(* IEC 61131-3 sources: teller/JD_Teller_LC2_V11/Class/SafetyManager (part 3) *)

            exit;
          end_if;

          pHelpManaging := pHelpManaging^.pNext;
        end_while;
      end_if;

      pHelpPdo := pHelpPdo^.pNext;
    end_while;

    pHelpConfig := pHelpConfig^.pNext;
  end_while;

END_FUNCTION

FUNCTION VIRTUAL SafetyManager::GetThisViaServerName
	VAR_INPUT
		pObjectDotServer 	: ^CHAR;
	END_VAR
	VAR_OUTPUT
		ThisPtr 	: pVoid;
	END_VAR
  VAR
    ChannelMode : CHMODE;
  END_VAR

  ThisPtr := NIL;

  if pObjectDotServer = NIL then
    return;
  end_if;

  // get thispointer to server via name
  ChannelMode := _LookUpEmbed_C(pObjectDotServer, #ThisPtr, NIL);

  // check if it's a server
  case ChannelMode of
    _CH_CMD,
    _CH_SVR:

  else
    ThisPtr := NIL;
    LogError(e_msg:="(SafetyManager::GetThisViaServerName) Couldn't get thispointer of server:");
    LogError(e_msg:=pObjectDotServer);
  end_case;

END_FUNCTION

FUNCTION SafetyManager::GetNewMovDO
	VAR_OUTPUT
		Index 	: INT;
	END_VAR
//  VAR
//  	sd_retval : DINT;
//  END_VAR

  Index := -1;

  if CopyCmdsUsed < MAX_PDO_COPY_CMDS then
    // check if there is one available but not used
    if CopyCmdsUsed < CopyCmdsAvailable then
      Index := CopyCmdsUsed;
      CopyCmdsUsed += 1;
    else
      // we have to create a new one

(*
// connection to varan manager required
      // add data object to copy our data
      sd_retval := pVaranManager^.AddMovDO(ud_dol_type:=VARAN_DOL_ISO
                                         , p_ud_handle:=(#aCopyCmds[CopyCmdsAvailable].pHandle)$^UDINT
                                         , p_ud_MovSettings:=( #aCopyCmds[CopyCmdsAvailable].pSettings)$^UDINT
                                         , ud_type := VM_PRIORITY_2
                                         );

      //look for an error
      if ( sd_retval <> 0 ) then
        ClassState := -9;
        LogError("(SafetyManager::GetNewMovDO) Failed to add a new copy command to the VaranManager!");
        return;
      end_if;
*)
      aCopyCmds[CopyCmdsAvailable].b_Ready4Action := FALSE;

      Index := CopyCmdsAvailable;

      CopyCmdsAvailable += 1;
      CopyCmdsUsed += 1;
    end_if;
  else
    LogError("Maximum of possible PDO copy commands reached!");
  end_if;

END_FUNCTION

FUNCTION SafetyManager::CheckCPUConfigs
	VAR_OUTPUT
		ConfigsOK 	: BOOL;
	END_VAR
  VAR
  	pHelpManaging   : ^t_ManagingComponent;
    pSourceManaging : ^t_ManagingComponent;
    pHelpConfig     : ^t_CfgListElem;
    pHelpPdo        : ^t_PdoListElem;
    pLastPdo        : ^t_PdoListElem;
    IsSource        : DINT;
    PDOCount : UDINT;
  END_VAR

  // before we go into the usual check routine, we have to ensure that we have enough virtual PDOs for writing interface frames (config holds a broadcast and we have to look for possible target modules)
  CreateVirtualPDOs();

  // initialize with true (normal case is that everything is ok => now we check for errors)
  ConfigsOK := TRUE;

  PDOCount := 0;

  // check if all non-optional modules are available and all corresponding domain managing module are synchron (if necessary)
  pHelpConfig := pConfigs;
  while pHelpConfig do
    pLastPdo := NIL;
    pHelpPdo := pHelpConfig^.pFirstPdoCfg;
    while pHelpPdo do
      // if it's an interface frame and no broadcast frame
      if pHelpPdo^.PdoInfo.Info.IsInterfacePDO then
        if (pHelpPdo^.PdoInfo.Info.IFBroadCast = FALSE) then

          // check if we have already added the domain interface to the IF List
          IsSource := -1; // -1 = not found, 0 = destination, 1 = source
          pSourceManaging := NIL;
          pHelpManaging := pFirstManagingInterfaceComponent;
          while pHelpManaging do
            // if source or destination of the PDO matches our managing module path => it's an interface frame to/from this domain
            if (To_StdLib.MemCmp(pHelpManaging^.pModulePath, pHelpPdo^.PdoInfo.pSourcePath, pHelpPdo^.PdoInfo.SourcePathLen) = 0) then
              pSourceManaging := pHelpManaging;
              IsSource := 1;
              exit;
            elsif (To_StdLib.MemCmp(pHelpManaging^.pModulePath, pHelpPdo^.PdoInfo.pDestPath, pHelpPdo^.PdoInfo.DestPathLen) = 0) then
              IsSource := 0;
              exit;
            end_if;

            pHelpManaging := pHelpManaging^.pNext;
          end_while;

          // if we got a source managing module and it isn't synchron
          if pSourceManaging then
            // if this pdo is not optional => the source module also isn't
            if pHelpPdo^.PdoInfo.Info.IsOptional = FALSE then
              pSourceManaging^.InfoBits.IsOptional := FALSE;
            end_if;

            if (pSourceManaging^.InfoBits.IsSynchron = FALSE) then
              if pHelpPdo^.PdoInfo.Info.IsOptional then
                // ignore it
  //              LogError("Info: Optional interface frame can't be received, because source domain is not connected or not synchron");

                // remove the PDO from the list (if not the receiver module would wait endless for the PDO and we can't send the set bus ready to quit errors of local PDOs)
                if pLastPdo then
                  // if we had already a PDO before in this configuration we have to skip the removed PDO with the next pointer
                  pLastPdo^.pNext := pHelpPdo^.pNext;

                  To_StdLib.Free(pHelpPdo^.PdoInfo.pSourcePath);
                  To_StdLib.Free(pHelpPdo^.PdoInfo.pDestPath);
                  To_StdLib.Free(pHelpPdo);

                  pHelpPdo := pLastPdo;
                else
                  // if it was the first PDO, we have to correct the first pointer
                  pHelpConfig^.pFirstPdoCfg := pHelpPdo^.pNext;

                  To_StdLib.Free(pHelpPdo^.PdoInfo.pSourcePath);
                  To_StdLib.Free(pHelpPdo^.PdoInfo.pDestPath);
                  To_StdLib.Free(pHelpPdo);

                  pHelpPdo := pHelpConfig^.pFirstPdoCfg;
                end_if;

                if pHelpPdo = NIL then
                  exit;
                end_if;
              else
                // non-optional interface frame domain missing => error
                LogError("ERROR! Non-Optional interface frame can't be received, because domain is not connected");
                ConfigsOK := FALSE;
                ClassState := -10;
              end_if;
            end_if;
          end_if;
        end_if;
      end_if;

      PDOCount += 1;

      pLastPdo := pHelpPdo;
      pHelpPdo := pHelpPdo^.pNext;
    end_while;

    pHelpConfig := pHelpConfig^.pNext;
  end_while;

  // if now PDOs found => reset the act ID to show that there are none
  if PDOCount = 0 then
    ActPDO_ID := 0;
  end_if;

END_FUNCTION

FUNCTION SafetyManager::RemoveLocalCPUCfg
	VAR_INPUT
		SafetyNumber 	: HDINT;
	END_VAR
  VAR
  	pHelpCfg    : ^t_LocalCfgListElem;
    i : UDINT;
  END_VAR

  if LocalCPUCfgNo then
    pHelpCfg := pFirstLocalCPUCfg;
    for i := 0 to (LocalCPUCfgNo-1) do
      if pHelpCfg^.SafetyNbr = SafetyNumber then
        // found it => deactivate it
        pHelpCfg^.ConfigSize := 0;
        pHelpCfg^.ConfigSent2Master := FALSE;
        exit;
      end_if;

      pHelpCfg := pHelpCfg^.pNext;
    end_for;
  end_if;

END_FUNCTION

FUNCTION SafetyManager::ClearRoutingInformations
  VAR
  	MyPara : CmdStruct;
    MyResult : results;
    pHelpManaging : ^t_ManagingComponent;
    i : UDINT;
    pHelpCfg      : ^t_LocalCfgListElem;
  END_VAR

  // we're flushin our stuff here

  // reset number of memorized safe cpu numbers
  SafeCPU_Nbr_No := 0;

  // set ID to zero for the next mapping assignment
  ActPDO_ID := 0;

  // reset interface frameno
  InterfaceFrameNo := 0;

  // reset local interface frameno
  LocalIFNo := 0;

  // clear configurations of safety-cpus
  FreeCfgLists();

  // clear number of copy DOs used
  CopyCmdsUsed := 0;

  // reset memory usage for isochronous transfer (the values are set when distributing the PDOs)
  MyPara.aPara[0] := 0;
  pHelpManaging := pFirstManagingInterfaceComponent;
  while pHelpManaging do
    pHelpManaging^.PDOReadMemUsed := 0;
    pHelpManaging^.PDOWriteMemUsed := 0;

    MyPara.uiCmd := CMD_SM_PDO_MEM_USAGE_WR;
    pHelpManaging^.pThis^.NewInst(#MyPara, #MyResult);

    MyPara.uiCmd := CMD_SM_PDO_MEM_USAGE_RD;
    pHelpManaging^.pThis^.NewInst(#MyPara, #MyResult);

    pHelpManaging^.InfoBits.HasBeenFlushed      := FALSE;
    pHelpManaging^.InfoBits.NewTimeSyncPossible := FALSE;
    pHelpManaging^.InfoBits.SubDomainsSynchron  := FALSE;
    pHelpManaging^.InfoBits.GotIFInfo           := FALSE;
    pHelpManaging^.InfoBits.LocalConfigReady    := FALSE;
    pHelpManaging^.InfoBits.IsOptional          := TRUE;  // initialize with true, later in the init process (CheckCPUConfigs) it's checked and corrected if necessary
    // synchron bit is already true at this time (or the timeout has expired)

    pHelpManaging^.DomainNr := 16#FF;

    pHelpManaging^.SubDomainsUsed := 0;
    _memset(dest:=#pHelpManaging^.SubDomainNr, usByte:=16#FF, cntr:=sizeof(pHelpManaging^.SubDomainNr));

    pHelpManaging^.ModuleNo := 0;
    _memset(dest:=#pHelpManaging^.ModuleInfo, usByte:=16#00, cntr:=sizeof(pHelpManaging^.ModuleInfo));

    pHelpManaging := pHelpManaging^.pNext;
  end_while;

  // all local cpu configs have to be sent again on reconnect
  if LocalCPUCfgNo then
    pHelpCfg := pFirstLocalCPUCfg;
    for i := 0 to (LocalCPUCfgNo-1) do
      pHelpCfg^.ConfigSent2Master := FALSE;

      pHelpCfg := pHelpCfg^.pNext;
    end_for;
  end_if;

END_FUNCTION

FUNCTION SafetyManager::CheckPDORecycle
	VAR_INPUT
		SourceDest 	: t_SourceDest;
		pNewPDO 	: ^t_PDOElement;
	END_VAR
	VAR_OUTPUT
		pRecyclePDO 	: ^t_PDOElement;
	END_VAR
  VAR
  	i : UDINT;
    pHelpInfo : ^t_PDOModuleInfo;
    pSearchInfo : ^t_PDOModuleInfo;
    ppHelpManaging : ^t_pManagingComponent;
    pSearchManaging : ^t_ManagingComponent;
  END_VAR

  // initialize with invalid
  pRecyclePDO := NIL;

  // if we have no pdoelements yet, quit
  if PDOElementNo = 0 then
    return;
  end_if;

  // we search for a PDO with the same source (then it contains the same data)
  pHelpInfo := #aPDOElements[0].SourceInfo;
  pSearchInfo := #pNewPDO^.SourceInfo;

  case SourceDest of
    SourceDest_IsSource:
      ppHelpManaging := #aPDOElements[0].pManagingSource;
      pSearchManaging := pNewPDO^.pManagingSource;
    SourceDest_IsDest:
      ppHelpManaging := #aPDOElements[0].pManagingDest;
      pSearchManaging := pNewPDO^.pManagingDest;
  else
    return;
  end_case;

  // check if we already have the path info of this source/destination
  for i := 0 to (PDOElementNo-1) do
    // if managing node, pathlength and path matches
    if (ppHelpManaging^ = pSearchManaging) & (pHelpInfo^.PathLen = pSearchInfo^.PathLen) & (To_StdLib.MemCmp(pHelpInfo^.pPath, pSearchInfo^.pPath, pHelpInfo^.PathLen) = 0) then
      // we found our PDO to recycle (PDO is already tranferred over this managing node
      pRecyclePDO := #aPDOElements[i];
      return;
    end_if;

    pHelpInfo       += sizeof(t_PDOElement);
    ppHelpManaging  += sizeof(t_PDOElement);
  end_for;

END_FUNCTION

FUNCTION SafetyManager::AddManagingInfo
	VAR_INPUT
		pPara 	: ^CmdStruct;
	END_VAR
  VAR
  	pHelpManaging : ^t_ManagingComponent;
  END_VAR

(*
  Parameter description:
  0..pointer to write PDOs in VARAN manager DPRAM
  1..pointer to read PDOs in VARAN manager DPRAM
  2..thispointer of calling class
  3..pointer to write PDOs in internal memory
  4..pointer to read PDOs in internal memory
  5..maximum available space for write PDOs in bytes
  6..maximum available space for read PDOs in bytes
*)

  pHelpManaging := pFirstManagingInterfaceComponent;
  while pHelpManaging do
    if pHelpManaging^.pThis = pPara^.aPara[2]$pVirtualBase then
      exit;
    end_if;

    pHelpManaging := pHelpManaging^.pNext;
  end_while;

  if pHelpManaging then
    pHelpManaging^.pPDOWriteSpaceDPRAM  := pPara^.aPara[0]$^USINT;
    pHelpManaging^.pPDOReadSpaceDPRAM   := pPara^.aPara[1]$^USINT;

    pHelpManaging^.pPDOWriteSpace       := pPara^.aPara[3]$^USINT;
    pHelpManaging^.pPDOReadSpace        := pPara^.aPara[4]$^USINT;

    pHelpManaging^.PDOWriteMemAvailable := pPara^.aPara[5]$UDINT;
    pHelpManaging^.PDOReadMemAvailable  := pPara^.aPara[6]$UDINT;

    pHelpManaging^.ud_HandlePDOWriteSpaceDPRAM  := pPara^.aPara[7]$UDINT;
    pHelpManaging^.ud_HandlePDOReadSpaceDPRAM   := pPara^.aPara[8]$UDINT;

  end_if;

END_FUNCTION

FUNCTION SafetyManager::CheckModuleUsage
	VAR_INPUT
		Length 	: UINT;
		pData 	: ^void;
	END_VAR
	VAR_OUTPUT
		retcode 	: DINT;
	END_VAR
  VAR
    pDataHelp : ^void;
    i : UDINT;
    TmpPathLen : UINT;
    TempCfgNo : USINT;
    ModuleCfgInfo : t_ModuleCfgInfo;
    PdoCfgInfo : t_PdoCfgInfo;
  END_VAR

(*
    Memory structure:
      4 Byte: SafetyNumber of CPU (is already there from initialisation in CSCP011_IM::InitSafeModule)
      1 Byte: Number of module configurations which are following
      for every module configuration (first is always the CPU itself)
        1 Byte: Info
        4 Byte: Interface Frame Source SafetyNumber (0 if it is no source for interface frames)
        4 Byte: Interface Frame CRC
        1 Byte: Number of destination inferface frame CRCs
        x Byte: Destination interface frame CRCs (number * sizeof(HDINT)
        2 Byte: Length of hardware path
        x Byte (depending on length in the 2 byte before): Hardwarepath
        2 Byte: Length of compressed hardware path
        x Byte (depending on length in the 2 byte before): Compressed Hardwarepath
        1 Byte: PDO out length for this module
      1 Byte: Number of pdo configurations which are following
      for every PDO configuration
        1 Byte: PDO length
        1 Byte: Interface frame info
        4 Byte: Interface CRC
        2 Byte: Length of source hardware path
        x Byte (depending on length in the 2 byte before): Hardwarepath of source
        2 Byte: Length of destination hardware path
        x Byte (depending on length in the 2 byte before): Hardwarepath of destination
      1 Byte: Number of slave configurations which are following
      for every slave configuration
        1 Byte: Info
        4 Byte: InterfaceCRC
        2 Byte: Length of hardware path
        x Byte (depending on length in the 2 byte before): Hardwarepath
        2 Byte: Length of compressed hardware path
        x Byte (depending on length in the 2 byte before): Compressed Hardwarepath
*)

  // check if the configuration is valid (pData <> NIL) & (Length must be at least 4 byte for SafetyNbr + 1 byte module cfg number + 1 byte pdo cfg number + 1 byte slave cfc number)
  if pData & (Length >= 7)  then

    retcode := 0;

    pDataHelp := pData;

    // skip safety number of the safety cpu
    pDataHelp += sizeof(HDINT);

    // number of module configurations which follow now
    TempCfgNo := pDataHelp^$USINT;

    // skip number of module configurations
    pDataHelp += sizeof(USINT);

    // module configurations
    if TempCfgNo then
      for i := 0 to (TempCfgNo-1) do
        // info
        ModuleCfgInfo := pDataHelp^$t_ModuleCfgInfo;

        // skip info
        pDataHelp += sizeof(BSINT);

        // skip safety number of interface frame source
        pDataHelp += sizeof(HDINT);

        // skip interface CRC of interface frame
        pDataHelp += sizeof(HDINT);

        // interface frame destination CRCs
        if ModuleCfgInfo.IsInterfaceDest then
          // number of CRCs
          TmpPathLen := pDataHelp^$USINT;

          // skip number of CRCs
          pDataHelp += sizeof(USINT);

          // skip interface destination CRCs
          pDataHelp += TmpPathLen * sizeof(HDINT);
        end_if;

        // length of hardware path
        TmpPathLen := pDataHelp^$UINT;

        // skip length of hardware path
        pDataHelp += sizeof(UINT);

        SetModuleUsed(PathLen:=TmpPathLen, pPath:=pDataHelp$^USINT, IgnoreOptional:=FALSE, IsOptional:=ModuleCfgInfo.IsOptional, IsInterfaceDomain := FALSE);

        // skip hardware path
        pDataHelp += TmpPathLen;

        // length of compressed hardware path
        TmpPathLen := pDataHelp^$UINT; // save some time with this local variable

        // skip length of compressed hardware path
        pDataHelp += sizeof(UINT);

        // skip compressed hardware path
        pDataHelp += TmpPathLen;

        // skip pdo out length of this module
        pDataHelp += sizeof(USINT);
      end_for;
    end_if;

    // number of Pdo configurations which follow now
    TempCfgNo := pDataHelp^$USINT;

    // skip number of pdo configurations
    pDataHelp += sizeof(USINT);

    // Pdo configurations
    if TempCfgNo then
      for i := 0 to (TempCfgNo-1) do
        // skip pdo length
        pDataHelp += sizeof(USINT);

        // is it an interface pdo?
        PdoCfgInfo := pDataHelp^$t_PdoCfgInfo;

        // skip info
        pDataHelp += sizeof(BSINT);

        // skip interface CRC
        pDataHelp += sizeof(HDINT);

        // length of source hardware path
        TmpPathLen := pDataHelp^$UINT;

        // skip length of source hardware path
        pDataHelp += sizeof(UINT);

        SetModuleUsed(PathLen:=TmpPathLen, pPath:=pDataHelp$^USINT, IgnoreOptional:=FALSE, IsOptional:=PdoCfgInfo.IsOptional, IsInterfaceDomain := PdoCfgInfo.IsInterfacePDO);

        // skip source hardware path
        pDataHelp += TmpPathLen;

        // length of destination hardware path
        TmpPathLen := pDataHelp^$UINT;

        // skip length of destination hardware path
        pDataHelp += sizeof(UINT);

        // a destination module doesn't influence the optional property=> ignore the optional setting
        SetModuleUsed(PathLen:=TmpPathLen, pPath:=pDataHelp$^USINT, IgnoreOptional:=TRUE, IsOptional:=FALSE, IsInterfaceDomain := PdoCfgInfo.IsInterfacePDO);

        // skip destination hardware path
        pDataHelp += TmpPathLen;
      end_for;
    end_if;

    // number of slave configurations which follow now
    TempCfgNo := pDataHelp^$USINT;

    // skip number of slave configurations
    pDataHelp += sizeof(USINT);

    // slave configurations
    if TempCfgNo then
      for i := 0 to (TempCfgNo-1) do
        // skip info
        pDataHelp += sizeof(BSINT);

        // skip InterfaceCRC
        pDataHelp += sizeof(HDINT);

        // length of hardwarepath
        TmpPathLen := pDataHelp^$UINT; // save some time with this local variable

        // skip length of hardwarepath
        pDataHelp += sizeof(UINT);

        // skip hardwarepath
        pDataHelp += TmpPathLen;

        // length of compressed hardwarepath
        TmpPathLen := pDataHelp^$UINT; // save some time with this local variable

        // skip length of compressed hardwarepath
        pDataHelp += sizeof(UINT);

        // skip compressed hardwarepath
        pDataHelp += TmpPathLen;
      end_for;
    end_if;

    // check if the given size matches the memory structure
    if (pDataHelp$UDINT - pData$UDINT) <> Length then
      LogError("(SafetyManager::CheckModuleUsage) Invalid configuration data given (length doesn't match memory structure)");
      retcode := -3;
      return;
    end_if;
  else
    // invalid configuration
    LogError("(SafetyManager::CheckModuleUsage) Found invalid safety cpu configuration: Pointer or size wrong");
    retcode := -1;
  end_if;

END_FUNCTION

FUNCTION SafetyManager::SetModuleUsed
	VAR_INPUT
		PathLen 	: UINT;
		pPath 	: ^USINT;
		IgnoreOptional 	: BOOL;
		IsOptional 	: BOOL;
		IsInterfaceDomain 	: BOOL;
	END_VAR
  VAR
    pHelpManaging : ^t_ManagingComponent;
    pHelpSafety : ^t_SafetyComponent;
    TempPath : ARRAY [0..99] OF USINT;
  END_VAR

  // search for the hardware path

  // start with the safety components
  pHelpSafety := pFirstSafetyComponent;
  while pHelpSafety & pHelpSafety^.pPath do
    // we have 1 byte path length on the safety component but we got a 2 byte path length from the configuration
    // furthermore the pPath string could be over more domains and we have only our local path => check if length is bigger and if there is a domain escape right before the domain number
    if ((pPath^ = pHelpSafety^.pPath^) | ((pPath^ > pHelpSafety^.pPath^) & ((pPath + 1 + pPath^ - pHelpSafety^.pPath^)^ = HWT_ESCAPE_DOMAIN))) &
       (To_StdLib.MemCmp(pHelpSafety^.pPath + 1, pPath + 2 + pPath^ - pHelpSafety^.pPath^, pHelpSafety^.pPath^) = 0) then
      // only set IsOptional to false (has been initialized with true)
      if (IsOptional = FALSE) & (IgnoreOptional = FALSE) then
        pHelpSafety^.InfoBits.IsOptional := FALSE;
      end_if;
      return;
    end_if;

    pHelpSafety := pHelpSafety^.pNext;
  end_while;

  // if not found, continue with the managing interface components
  pHelpManaging := pFirstManagingInterfaceComponent;
  while pHelpManaging do
    if (To_StdLib.MemCmp(pHelpManaging^.pModulePath, pPath, PathLen) = 0) then
      // only set IsOptional to false (has been initialized with true)
      if (IsOptional = FALSE) & (IgnoreOptional = FALSE) then
        pHelpManaging^.InfoBits.IsOptional := FALSE;
      end_if;
      return;
    end_if;

    pHelpManaging := pHelpManaging^.pNext;
  end_while;

  _memcpy(ptr1:=#TempPath[0], ptr2:=pPath, cntr:=PathLen$USINT);

END_FUNCTION

FUNCTION SafetyManager::CreateTimeSyncList
  VAR
  	pHelp : ^t_TimeSyncElement;
  	pHelpSafety   : ^t_SafetyComponent;
  	pHelpManaging : ^t_ManagingComponent;
  END_VAR

  // first we stop time syncing (if active) to prevent crashing due tue a running time synchronisation
  pActTimeSyncElement := NIL;

  // if there is an old list, free it first
  if pFirstTimeSyncElement then
    // open the ring (set the next pointer of the last element to NIL)
    pFirstTimeSyncElement^.pPrev^.pNext := NIL;

    // remove the elements
    while pFirstTimeSyncElement do
      pHelp := pFirstTimeSyncElement;
      pFirstTimeSyncElement := pFirstTimeSyncElement^.pNext;

      To_StdLib.Free(mptr:=pHelp);
    end_while;
  end_if;

  pHelpSafety := pFirstSafetyComponent;
  while pHelpSafety do
    // if it's a module with not only inputs (then there's nothing to synchronize with) => trigger it for time synchronisation
    if (pHelpSafety^.InfoBits.OnlyInputs = FALSE) then
      AddTimeSyncElement(pManaging:=NIL, pSafety:=pHelpSafety, IsInterfaceDomain := FALSE);
    end_if;

    pHelpSafety := pHelpSafety^.pNext;
  end_while;

  // interface domains will not get our token, they got their own
  pHelpManaging := pFirstManagingInterfaceComponent;
  while pHelpManaging do
    AddTimeSyncElement(pManaging:=pHelpManaging, pSafety:=NIL, IsInterfaceDomain := TRUE);

    pHelpManaging := pHelpManaging^.pNext;
  end_while;

END_FUNCTION

FUNCTION SafetyManager::AddTimeSyncElement
	VAR_INPUT
		pManaging 	: ^t_ManagingComponent;
		pSafety 	: ^t_SafetyComponent;
		IsInterfaceDomain 	: BOOL;
	END_VAR
  VAR
    pLast : ^t_TimeSyncElement;
  	pHelp : ^t_TimeSyncElement;
  END_VAR

  // first we have to allocate some memory for the new element
  if pFirstTimeSyncElement = NIL then
    pFirstTimeSyncElement$pVoid := To_StdLib.Malloc(size:=sizeof(t_TimeSyncElement));
    pLast := pHelp := pFirstTimeSyncElement;
  else
    // check if we got this already
    pHelp := pFirstTimeSyncElement;
    repeat
      if pSafety & (pHelp^.pSafety = pSafety) then
        // already in list => leave
        return;
      end_if;

      if pManaging & (pHelp^.pManaging = pManaging) then
        // already in list => leave
        return;
      end_if;

      pHelp := pHelp^.pNext;
    until (pHelp = pFirstTimeSyncElement) end_repeat;

    pHelp$pVoid := To_StdLib.Malloc(size:=sizeof(t_TimeSyncElement));
    pLast := pFirstTimeSyncElement^.pPrev;
  end_if;

  if pHelp then
    // close the double linked ring with the new elements
    pFirstTimeSyncElement^.pPrev := pHelp;
    pHelp^.pNext := pFirstTimeSyncElement;

    pHelp^.pPrev := pLast;
    pLast^.pNext := pHelp;

    pHelp^.InfoBits := 0;
    pHelp^.InfoBits.IsInterfaceDomain := IsInterfaceDomain;

    pHelp^.pManaging := pManaging;
    pHelp^.pSafety   := pSafety;

    // managing modules
    if (pManaging <> NIL) then
      pHelp^.InfoBits.IsManagingModule := TRUE;
      pHelp^.pThis := pManaging^.pThis;

      // if it's the master connection
      if pManaging^.InfoBits.IsConnectionToMaster then
        // remember it
        pHelp^.InfoBits.IsConnectionToMaster := TRUE;

        // and make it the end of the list
        pFirstTimeSyncElement := pHelp^.pNext;

        // remember that we got a master connection
        pMasterTimeSyncElement := pHelp;

      elsif pMasterTimeSyncElement then
        // if we're not master and there is already a master time sync element in the list, we have to make it the last element
        pFirstTimeSyncElement := pMasterTimeSyncElement^.pNext;
      end_if;
    else
      // safety modules
      pHelp^.InfoBits.IsManagingModule := FALSE;
      pHelp^.pThis := pSafety^.pThis;

    // insert new safety modules at the beginning (managing modules at the end)
      pFirstTimeSyncElement := pHelp;
    end_if;

  else
    ClassState := -1;
    LogError("(SafetyManager::AddTimeSyncElement) Failed to allocate memory for a new Element");
  end_if;

END_FUNCTION

FUNCTION SafetyManager::CreateVirtualPDOs
  VAR
  	pHelpManaging   : ^t_ManagingComponent;
    pHelpConfig     : ^t_CfgListElem;
    pHelpPdo        : ^t_PdoListElem;
    TempPDO         : t_PdoCfg;
    pSearchConfig   : ^t_CfgListElem;
    pSearchPdo      : ^t_PdoListElem;
  END_VAR

  pHelpConfig := pConfigs;
  while pHelpConfig do
    pHelpPdo := pHelpConfig^.pFirstPdoCfg;
    while pHelpPdo do
      // check if it's a broadcast
      if (pHelpPdo^.PdoInfo.Info.IFBroadCast) & (pHelpPdo^.PdoInfo.Info.VirtualPDOsCreated = FALSE) then
        // found one => create virtual PDOs from it (add them to the same configuration)

        // prepare new virtual PDO
        TempPDO := pHelpPdo^.PdoInfo;

        TempPDO.Info.IFBroadCast := FALSE;
        TempPDO.Info.VirtualPDO := TRUE;

        // add a new PDO for every interface managing module
        pHelpManaging := pFirstManagingInterfaceComponent;
        while pHelpManaging do
          // change destination path to the actual module
          TempPDO.DestPathLen := pHelpManaging^.pModulePath^ + 2;
          TempPDO.pDestPath := pHelpManaging^.pModulePath;

          if AddVirtualPDOToCfg(pCfg:=pHelpConfig, pNewPDO:=#TempPDO) then
            LogError(e_msg:="(SafetyManager::CreateVirtualPDOs) Failed to allocate memory for a new virtual PDO");
          end_if;

          pHelpManaging := pHelpManaging^.pNext;
        end_while;

        // search in all configs (if there are other) for a pdo with this interface CRC as source
        pSearchConfig := pConfigs;
        while pSearchConfig do
          pSearchPdo := pSearchConfig^.pFirstPdoCfg;
          while pSearchPdo do
            // we must not manipulate our help pdo
            if pSearchPdo <> pHelpPdo then
              // check if the interface CRC appears in any PDO
              if pSearchPdo^.PdoInfo.InterfaceCRC = pHelpPdo^.PdoInfo.InterfaceCRC then
                // now take the source path of the broadcast PDO and use it as source path for this PDO
                To_StdLib.Free(mptr:=pSearchPdo^.PdoInfo.pSourcePath);

                pSearchPdo^.PdoInfo.pSourcePath$pVoid := To_StdLib.Malloc(size:=pHelpPdo^.PdoInfo.SourcePathLen);

                // save source hardwarepath
                if pSearchPdo^.PdoInfo.pSourcePath then
                  _memcpy(ptr1:=pSearchPdo^.PdoInfo.pSourcePath, ptr2:=pHelpPdo^.PdoInfo.pSourcePath, cntr:=pHelpPdo^.PdoInfo.SourcePathLen);
                  pSearchPdo^.PdoInfo.SourcePathLen := pHelpPdo^.PdoInfo.SourcePathLen;

                  // source and destination of this PDO are both local safe cpu modules which communicate with each other via interface frames => store them in extra list for routing SDOs and TDOs
                  AddToLocalIFs(#pSearchPdo^.PdoInfo);
                else
                  LogError(e_msg:="(SafetyManager::CreateVirtualPDOs) Failed to allocate memory for a source path");
                  pSearchPdo^.PdoInfo.SourcePathLen := 0;
                  ClassState := -1;
                end_if;
              end_if;
            end_if;

            pSearchPdo := pSearchPdo^.pNext;
          end_while;

          pSearchConfig := pSearchConfig^.pNext;
        end_while;
        pHelpPdo^.PdoInfo.Info.VirtualPDOsCreated := TRUE;
      end_if;

      pHelpPdo := pHelpPdo^.pNext;
    end_while;

    pHelpConfig := pHelpConfig^.pNext;
  end_while;

END_FUNCTION

FUNCTION SafetyManager::AddVirtualPDOToCfg
	VAR_INPUT
		pCfg 	: ^t_CfgListElem;
		pNewPDO 	: ^t_PdoCfg;
	END_VAR
	VAR_OUTPUT
		retcode 	: DINT;
	END_VAR
  VAR
    pHelpPdo        : ^t_PdoListElem;
    TempLen         : UINT;
  END_VAR

  retcode := 0;

  if pCfg^.pFirstPdoCfg = NIL then
    // first PDO in this cfg (should not be possible, because the template for this PDO is also in the same config)
    pCfg^.pFirstPdoCfg$pVoid := To_StdLib.Malloc(size:=sizeof(t_PdoListElem));
    pHelpPdo := pCfg^.pFirstPdoCfg;
  else
    // search a place for the new PDO
    pHelpPdo := pCfg^.pFirstPdoCfg;
    while pHelpPdo^.pNext do

      pHelpPdo := pHelpPdo^.pNext;
    end_while;

    pHelpPdo^.pNext$pvoid := To_StdLib.Malloc(size:=sizeof(t_PdoListElem));
    pHelpPdo := pHelpPdo^.pNext;
  end_if;

  if pHelpPdo then
    // init the values
    pHelpPdo^.PdoInfo.PdoLen        := pNewPDO^.PdoLen;
    pHelpPdo^.PdoInfo.Info          := pNewPDO^.Info;
    pHelpPdo^.PdoInfo.InterfaceCRC  := pNewPDO^.InterfaceCRC;

    // length of source hardwarepath
    TempLen := pNewPDO^.SourcePathLen; // save some time with this local variable
    pHelpPdo^.PdoInfo.SourcePathLen := TempLen;

    // allocate memory for the source module path
    pHelpPdo^.PdoInfo.pSourcePath$pVoid := To_StdLib.Malloc(size:=TempLen);
    if pHelpPdo^.PdoInfo.pSourcePath = NIL then
      ClassState := -1;
      retcode := -2;
      return;
    end_if;

    // save source hardwarepath
    _memcpy(ptr1:=pHelpPdo^.PdoInfo.pSourcePath, ptr2:=pNewPDO^.pSourcePath, cntr:=TempLen);

    // length of destination hardwarepath
    TempLen := pNewPDO^.DestPathLen; // save some time with this local variable
    pHelpPdo^.PdoInfo.DestPathLen := TempLen;

    // allocate memory for the destination module path
    pHelpPdo^.PdoInfo.pDestPath$pVoid := To_StdLib.Malloc(size:=TempLen);
    if pHelpPdo^.PdoInfo.pDestPath = NIL then
      ClassState := -1;
      retcode := -2;
      return;
    end_if;

    // save destination hardwarepath
    _memcpy(ptr1:=pHelpPdo^.PdoInfo.pDestPath, ptr2:=pNewPDO^.pDestPath, cntr:=TempLen);

    // now we give it an ID and increase the number for the next pdo
    pHelpPdo^.PdoInfo.PDO_ID := ActPDO_ID;
    ActPDO_ID += 1;

    pHelpPdo^.pNext                  := NIL;
  else
    ClassState := -1;
    retcode := -2;
    return;
  end_if;

END_FUNCTION

FUNCTION SafetyManager::AddToLocalIFs
	VAR_INPUT
		pHelpPDO 	: ^t_PdoCfg;
	END_VAR
  VAR
  	AddSource : BOOL;
    i : USINT;
    pHelpSafety : ^t_SafetyComponent;
  END_VAR

  // check if there is still room for new modules
  if LocalIFNo < MAX_INTERNAL_IF_MODULES then

    AddSource := TRUE;

    // if there is a list, check if any of our modules are already in the list
    if LocalIFNo then
      for i := 0 to (LocalIFNo-1) do
        // check if crc matches
        if (aLocalIFs[i].InterfaceCRC = pHelpPDO^.InterfaceCRC) then
          AddSource := FALSE;
          exit;
        end_if;
      end_for;
    end_if;

    // now we know how many we have to add to the list. if there are modules to add and there is enough space for all of them => do it
    if AddSource then
      // search it in the local modules
      pHelpSafety := pFirstSafetyComponent;
      while pHelpSafety do
        // if the path matches, add the module to the list

        // source module
        if (pHelpSafety^.PathLen = (pHelpPDO^.SourcePathLen - 1)) &
        // we compare the last x byte (where x is the length of the local path including the domain) because we got different length info sizes (1 byte vs. 2 byte)
           (To_StdLib.MemCmp(pHelpSafety^.pPath + 1, pHelpPDO^.pSourcePath + 2 + pHelpPDO^.pSourcePath^ - pHelpSafety^.pPath^, pHelpSafety^.pPath^) = 0) then
          aLocalIFs[LocalIFNo].InterfaceCRC  := pHelpPDO^.InterfaceCRC;
          aLocalIFs[LocalIFNo].pSafetyModule := pHelpSafety;
          LocalIFNo += 1;
          exit;
        end_if;

        pHelpSafety := pHelpSafety^.pNext;
      end_while;
    end_if;
  end_if;

END_FUNCTION

FUNCTION SafetyManager::IFInfoNotArrivedYet
	VAR_INPUT
		pThis 	: pVirtualBase;
	END_VAR
	VAR_OUTPUT
		InfoNotAvailable 	: BOOL;
	END_VAR
  VAR
  	pHelpManaging : ^t_ManagingComponent;
  END_VAR

	InfoNotAvailable := FALSE;

  pHelpManaging := pFirstManagingInterfaceComponent;
  while pHelpManaging do
    if pHelpManaging^.pThis = pThis then
      if pHelpManaging^.InfoBits.GotIFInfo = FALSE then
        InfoNotAvailable := TRUE;
      end_if;
      return;
    end_if;

    pHelpManaging := pHelpManaging^.pNext;
  end_while;

END_FUNCTION

#pragma warning(disable:74)
FUNCTION SafetyManager::StartTimeMeasurement
	VAR_INPUT
		usMode (EAX) 	: DINT;
	END_VAR
#ifdef VM_CLASS_TIME_MEASUREMENT
  VAR
  	tmpTime : ^t_TimeMeasurementVaran;
  END_VAR

  case usMode of

    //-----------------------------------------------------------

    VARANTIME_RT:
      tmpTime := #s_TimeRt;

    //-----------------------------------------------------------

    VARANTIME_RTPOSTSCAN:
      tmpTime := #s_TimeRtPostScan;

    //-----------------------------------------------------------

    VARANTIME_CY:
      tmpTime := #s_TimeCy;

    //-----------------------------------------------------------

  end_case;

  if ( tmpTime^.us_Activate ) then
//    Save_Flg();
//    CLI();
    tmpTime^.ud_Timemark := OS_READMICROSEC();
  end_if;

#endif

END_FUNCTION

FUNCTION SafetyManager::StopTimeMeasurement
	VAR_INPUT
		usMode (EAX) 	: DINT;
	END_VAR
#ifdef VM_CLASS_TIME_MEASUREMENT
  VAR
  	tmpTime : ^t_TimeMeasurementVaran;
  END_VAR

  case usMode of

    //-----------------------------------------------------------

    VARANTIME_RT:
      tmpTime := #s_TimeRt;

    //-----------------------------------------------------------

    VARANTIME_RTPOSTSCAN:
      tmpTime := #s_TimeRtPostScan;

    //-----------------------------------------------------------

    VARANTIME_CY:
      tmpTime := #s_TimeCy;

    //-----------------------------------------------------------

  end_case;

	if ( tmpTime^.us_Activate ) then

		//get actual time
		tmpTime^.ud_ActualTime := OS_READMICROSEC();
    tmpTime^.ud_ActualTime -= tmpTime^.ud_Timemark;

		//look for maximum time
		if ( tmpTime^.ud_ActualTime > tmpTime^.ud_MaximalTime ) then
			tmpTime^.ud_MaximalTime := tmpTime^.ud_ActualTime;
		end_if;

		//look for minimum time
		if ( tmpTime^.ud_ActualTime < tmpTime^.ud_MinimalTime ) then
			tmpTime^.ud_MinimalTime := tmpTime^.ud_ActualTime;
		end_if;

		//look for average time (100000 cycles)
		if ( tmpTime^.ud_AverageCounter = 100000 ) then

			tmpTime^.ud_AverageTime 	:= tmpTime^.ud_AverageSum / tmpTime^.ud_AverageCounter;
			tmpTime^.ud_AverageSum 	:= 0;
			tmpTime^.ud_AverageCounter := 0;

		else
			tmpTime^.ud_AverageSum += ( tmpTime^.ud_ActualTime / 100 );
			tmpTime^.ud_AverageCounter += 1;
		end_if;

//		STI();
//    Restore_Flg();
	end_if;

#endif

END_FUNCTION // Varan_Base::StopTimeMeasurement
#pragma warning(default:74)

FUNCTION SafetyManager::AnyIFDomainSynchron
	VAR_OUTPUT
		AnythingSynchron 	: BOOL;
	END_VAR
  VAR
    pHelpManaging   : ^t_ManagingComponent;
  END_VAR

  AnythingSynchron := FALSE;

  pHelpManaging := pFirstManagingInterfaceComponent;
  while pHelpManaging do
    if pHelpManaging^.InfoBits.IsSynchron then
      AnythingSynchron := TRUE;
      return;
    end_if;

    pHelpManaging := pHelpManaging^.pNext;
  end_while;

END_FUNCTION

FUNCTION SafetyManager::LocalIFsAvailable
	VAR_OUTPUT
		retcode 	: BOOL;
	END_VAR
  VAR
    pHelpCfg : ^t_CfgListElem;
    pHelpPdo : ^t_PdoListElem;
    pHelpModule : ^t_ModuleListElem;
  END_VAR

  retcode := FALSE;

  // add all local configs to our structure
  SendLocalCfgsToMaster();

  // check the local configs for interface frames
  pHelpCfg := pConfigs;
  while pHelpCfg do
    pHelpPdo := pHelpCfg^.pFirstPdoCfg;
    while pHelpPdo do
      if pHelpPdo^.PdoInfo.Info.IsInterfacePDO | pHelpPdo^.PdoInfo.Info.IFBroadCast then
        retcode := TRUE;
        return;
      end_if;

      pHelpPdo := pHelpPdo^.pNext;
    end_while;

    pHelpModule := pHelpCfg^.pFirstModuleCfg;
    while pHelpModule do
      if pHelpModule^.ModuleInfo.Info.IsInterfaceSource | pHelpModule^.ModuleInfo.Info.IsInterfaceDest then
        retcode := TRUE;
        return;
      end_if;

      pHelpModule := pHelpModule^.pNext;
    end_while;

    pHelpCfg := pHelpCfg^.pNext;
  end_while;

END_FUNCTION

FUNCTION SafetyManager::IsCPUModule
  VAR_INPUT
    ModuleType : t_e_ModuleType;
  END_VAR
  VAR_OUTPUT
  	retcode : BOOL;
  END_VAR

  case ModuleType of
    _CSCP01x,
    _SCP010,
    _SCP011:
      retcode := TRUE;
  else
    retcode := FALSE;
  end_case;

END_FUNCTION
